// TIA Portal V19 export
FUNCTION_BLOCK "HOT_SKIDS"   // FB19, LAD
{ S7_Optimized_Access := 'TRUE' }
// stored: MemoryReserve 100, SetENOAutomatically false
   VAR_INPUT
      TEMP_SP : Real;
      AUTO : Bool;
      START : Bool;
      STOP : Bool;
      PUMP_SEL_1 : Bool;
      PUMP_SEL_2 : Bool;
      PUMP_SEL_3 : Bool;
      EMG : Bool;
      FS_HE_OUTLET : Bool;
      MGLT_LSP : Real;
      HOLD_RESUME : Bool;
      TT01_fault : Bool;
      TT02_fault : Bool;
      TT03_fault : Bool;
      TT04_fault : Bool;
      MGLT_FAULT : Bool;
      HEADER_PRESSURE_SP : Real;
      MGLT_PV : Real;
      TEMP_PV : Real;
      HEADER_PRESSURE_PV : Real;
      "PUMP 1RPM" : Real;
      "PUMP 1 RPM_SP" : Real;
      "PUMP 2 RPM" : Real;
      "PUMP 2 RPM_SP" : Real;
      "PUMP 3 RPM" : Real;
      "PUMP 3 RPM_SP" : Real;
   END_VAR
   VAR_OUTPUT
      PUMP_1_CMD : Bool;
      PUMP_2_CMD : Bool;
      PUMP_3_CMD : Bool;
      RUNNING : Bool;
      HS_CV_CMD : Bool;
      PUMP_SEL : Int;
      PUMP_1_FAULTY : Bool;
      PUMP_2_FAULTY : Bool;
      PUMP_3_FAULTY : Bool;
   END_VAR
   VAR
      "STEP" : Int;
      IEC_Timer_0_Instance { S7_SetPoint := 'True'} : TP_TIME;
      ALL_OK : Bool;
      TRIG_1 : Bool;
      TRIG_2 : Bool;
      TRIG_3 : Bool;
      TRIG_4 : Bool;
      TRIG_5 : Bool;
      TRIG_6 : Bool;
      TRIG_7 : Bool;
      IEC_Timer_0_Instance_1 { S7_SetPoint := 'True'} : TP_TIME;
      IEC_Timer_0_Instance_2 { S7_SetPoint := 'True'} : TP_TIME;
   END_VAR
   VAR_TEMP   // added for the SCL form of the ladder/FBD networks
      _w1 : Bool;
      _w2 : Bool;
      _w3 : Bool;
      _w4 : Bool;
   END_VAR
BEGIN

REGION Network 1: PRECHECK
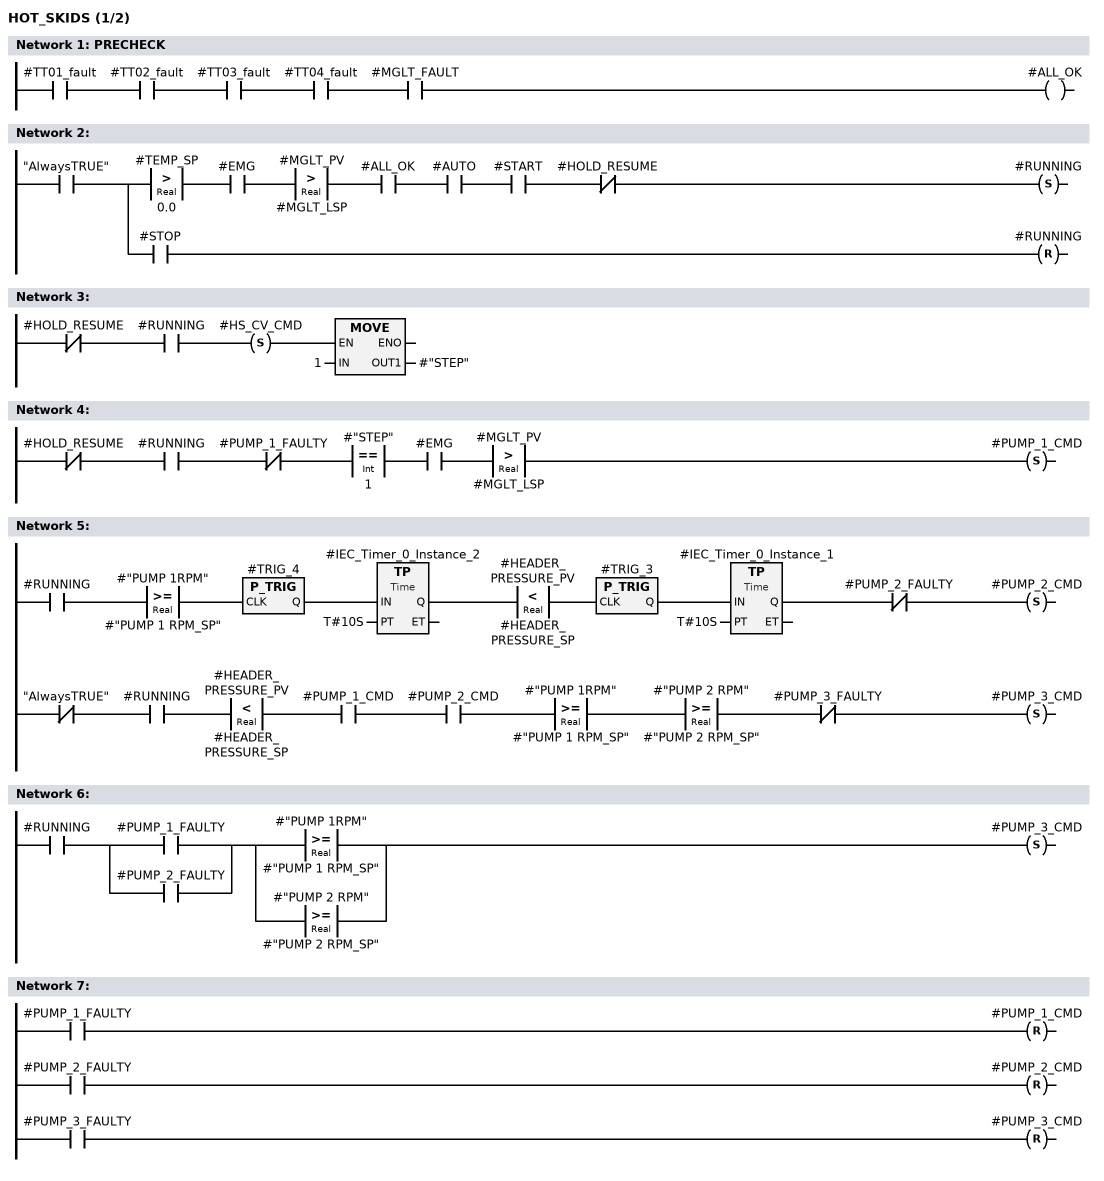
   RUNG wire#powerrail
      Contact( #TT01_fault )
      Contact( #TT02_fault )
      Contact( #TT03_fault )
      Contact( #TT04_fault )
      Contact( #MGLT_FAULT )
      Coil( #ALL_OK )
   END_RUNG
   // the same network as SCL:
   #ALL_OK := #TT01_fault AND #TT02_fault AND #TT03_fault AND #TT04_fault AND #MGLT_FAULT;
END_REGION

REGION Network 2
   RUNG wire#powerrail
      Contact( "AlwaysTRUE" )
      wire#w1
      { S7_Templates := "SrcType := Real" } GT_Contact(in1 := #TEMP_SP, in2 := 0.0)
      Contact( #EMG )
      { S7_Templates := "SrcType := Real" } GT_Contact(in1 := #MGLT_PV, in2 := #MGLT_LSP)
      Contact( #ALL_OK )
      Contact( #AUTO )
      Contact( #START )
      I_Contact( #HOLD_RESUME )
      S_Coil( #RUNNING )
   END_RUNG
   RUNG wire#w1
      Contact( #STOP )
      R_Coil( #RUNNING )
   END_RUNG
   // the same network as SCL:
   IF "AlwaysTRUE" AND (#TEMP_SP > 0.0) AND #EMG AND (#MGLT_PV > #MGLT_LSP) AND #ALL_OK AND #AUTO AND #START AND NOT #HOLD_RESUME THEN
       #RUNNING := TRUE;
   END_IF;
   IF "AlwaysTRUE" AND #STOP THEN #RUNNING := FALSE; END_IF;
END_REGION

REGION Network 3
   RUNG wire#powerrail
      I_Contact( #HOLD_RESUME )
      Contact( #RUNNING )
      S_Coil( #HS_CV_CMD )
      Move(in := 1, out1 => #"STEP")
   END_RUNG
   // the same network as SCL:
   IF NOT #HOLD_RESUME AND #RUNNING THEN
       #HS_CV_CMD := TRUE;
       #"STEP" := 1;
   END_IF;
END_REGION

REGION Network 4
   RUNG wire#powerrail
      I_Contact( #HOLD_RESUME )
      Contact( #RUNNING )
      I_Contact( #PUMP_1_FAULTY )
      { S7_Templates := "SrcType := Int" } EQ_Contact(in1 := #"STEP", in2 := 1)
      Contact( #EMG )
      { S7_Templates := "SrcType := Real" } GT_Contact(in1 := #MGLT_PV, in2 := #MGLT_LSP)
      S_Coil( #PUMP_1_CMD )
   END_RUNG
   // the same network as SCL:
   IF NOT #HOLD_RESUME AND #RUNNING AND NOT #PUMP_1_FAULTY AND (#"STEP" = 1) AND #EMG AND (#MGLT_PV > #MGLT_LSP) THEN
       #PUMP_1_CMD := TRUE;
   END_IF;
END_REGION

REGION Network 5
   RUNG wire#powerrail
      Contact( #RUNNING )
      { S7_Templates := "SrcType := Real" } GE_Contact(in1 := #"PUMP 1RPM", in2 := #"PUMP 1 RPM_SP")
      P_Trig( #TRIG_4 )
      { S7_Templates := "time_type := Time" } #IEC_Timer_0_Instance_2.TP(pt := T#10S, et =>)
      { S7_Templates := "SrcType := Real" } LT_Contact(in1 := #HEADER_PRESSURE_PV, in2 := #HEADER_PRESSURE_SP)
      P_Trig( #TRIG_3 )
      { S7_Templates := "time_type := Time" } #IEC_Timer_0_Instance_1.TP(pt := T#10S, et =>)
      I_Contact( #PUMP_2_FAULTY )
      S_Coil( #PUMP_2_CMD )
   END_RUNG
   RUNG wire#powerrail
      I_Contact( "AlwaysTRUE" )
      Contact( #RUNNING )
      { S7_Templates := "SrcType := Real" } LT_Contact(in1 := #HEADER_PRESSURE_PV, in2 := #HEADER_PRESSURE_SP)
      Contact( #PUMP_1_CMD )
      Contact( #PUMP_2_CMD )
      { S7_Templates := "SrcType := Real" } GE_Contact(in1 := #"PUMP 1RPM", in2 := #"PUMP 1 RPM_SP")
      { S7_Templates := "SrcType := Real" } GE_Contact(in1 := #"PUMP 2 RPM", in2 := #"PUMP 2 RPM_SP")
      I_Contact( #PUMP_3_FAULTY )
      S_Coil( #PUMP_3_CMD )
   END_RUNG
   // the same network as SCL:
   #_w1 := #RUNNING AND (#"PUMP 1RPM" >= #"PUMP 1 RPM_SP");
   #_w2 := #_w1 AND NOT #TRIG_4;   // rising edge
   #TRIG_4 := #_w1;
   #IEC_Timer_0_Instance_2(IN := #_w2, PT := T#10S);   // TP
   #_w3 := #IEC_Timer_0_Instance_2.Q AND (#HEADER_PRESSURE_PV < #HEADER_PRESSURE_SP);
   #_w4 := #_w3 AND NOT #TRIG_3;   // rising edge
   #TRIG_3 := #_w3;
   #IEC_Timer_0_Instance_1(IN := #_w4, PT := T#10S);   // TP
   IF #IEC_Timer_0_Instance_1.Q AND NOT #PUMP_2_FAULTY THEN #PUMP_2_CMD := TRUE; END_IF;
   IF NOT "AlwaysTRUE" AND #RUNNING AND (#HEADER_PRESSURE_PV < #HEADER_PRESSURE_SP) AND #PUMP_1_CMD AND #PUMP_2_CMD AND (#"PUMP 1RPM" >= #"PUMP 1 RPM_SP") AND (#"PUMP 2 RPM" >= #"PUMP 2 RPM_SP") AND NOT #PUMP_3_FAULTY THEN
       #PUMP_3_CMD := TRUE;
   END_IF;
END_REGION

REGION Network 6
   RUNG wire#powerrail
      Contact( #RUNNING )
      wire#w1
      Contact( #PUMP_1_FAULTY )
      wire#w2
      { S7_Templates := "SrcType := Real" } GE_Contact(in1 := #"PUMP 1RPM", in2 := #"PUMP 1 RPM_SP")
      wire#w3
      S_Coil( #PUMP_3_CMD )
   END_RUNG
   RUNG wire#w1
      Contact( #PUMP_2_FAULTY )
   END_RUNG wire#w2
   RUNG wire#w2
      { S7_Templates := "SrcType := Real" } GE_Contact(in1 := #"PUMP 2 RPM", in2 := #"PUMP 2 RPM_SP")
   END_RUNG wire#w3
   // the same network as SCL:
   IF #RUNNING AND (#PUMP_1_FAULTY OR #PUMP_2_FAULTY) AND ((#"PUMP 1RPM" >= #"PUMP 1 RPM_SP") OR (#"PUMP 2 RPM" >= #"PUMP 2 RPM_SP")) THEN
       #PUMP_3_CMD := TRUE;
   END_IF;
END_REGION

REGION Network 7
   RUNG wire#powerrail
      Contact( #PUMP_1_FAULTY )
      R_Coil( #PUMP_1_CMD )
   END_RUNG
   RUNG wire#powerrail
      Contact( #PUMP_2_FAULTY )
      R_Coil( #PUMP_2_CMD )
   END_RUNG
   RUNG wire#powerrail
      Contact( #PUMP_3_FAULTY )
      R_Coil( #PUMP_3_CMD )
   END_RUNG
   // the same network as SCL:
   IF #PUMP_1_FAULTY THEN #PUMP_1_CMD := FALSE; END_IF;
   IF #PUMP_2_FAULTY THEN #PUMP_2_CMD := FALSE; END_IF;
   IF #PUMP_3_FAULTY THEN #PUMP_3_CMD := FALSE; END_IF;
END_REGION

REGION Network 8
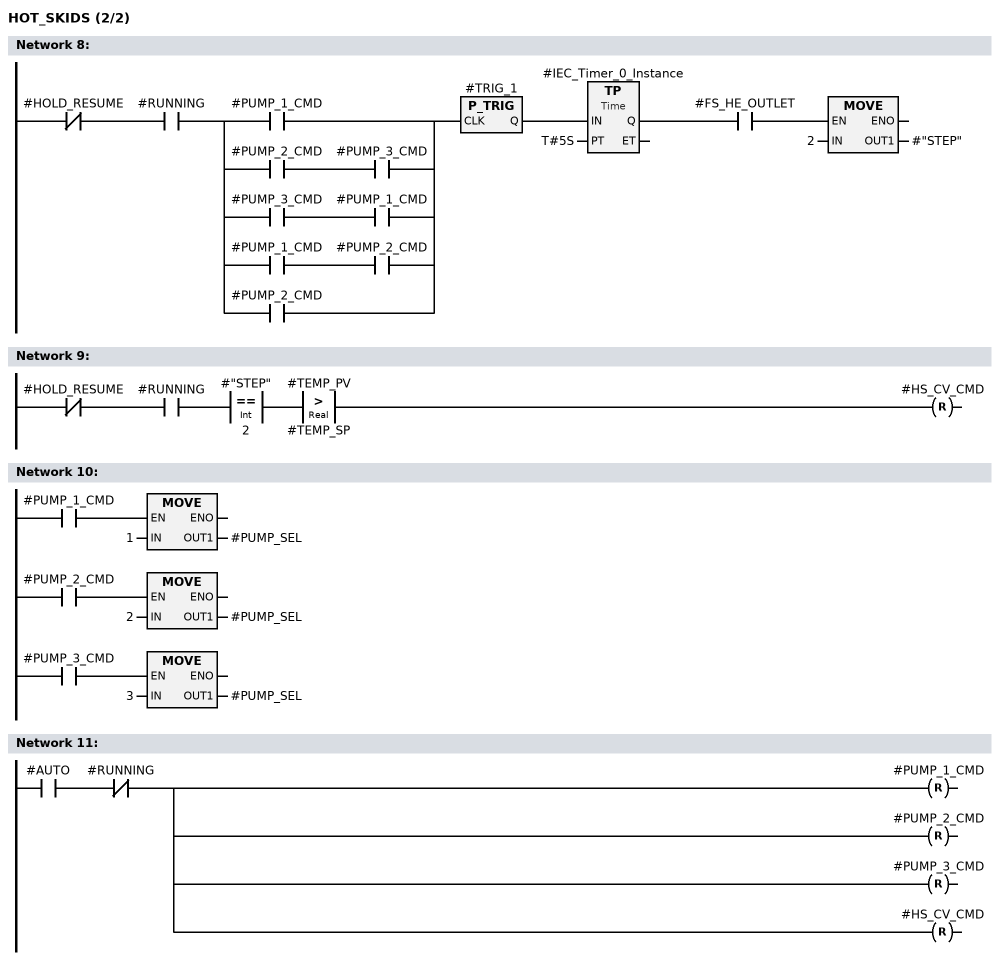
   RUNG wire#powerrail
      I_Contact( #HOLD_RESUME )
      Contact( #RUNNING )
      wire#w1
      Contact( #PUMP_1_CMD )
      wire#w2
      P_Trig( #TRIG_1 )
      { S7_Templates := "time_type := Time" } #IEC_Timer_0_Instance.TP(pt := T#5S, et =>)
      Contact( #FS_HE_OUTLET )
      Move(in := 2, out1 => #"STEP")
   END_RUNG
   RUNG wire#w1
      Contact( #PUMP_2_CMD )
      Contact( #PUMP_3_CMD )
   END_RUNG wire#w2
   RUNG wire#w1
      Contact( #PUMP_3_CMD )
      Contact( #PUMP_1_CMD )
   END_RUNG wire#w2
   RUNG wire#w1
      Contact( #PUMP_1_CMD )
      Contact( #PUMP_2_CMD )
   END_RUNG wire#w2
   RUNG wire#w1
      Contact( #PUMP_2_CMD )
   END_RUNG wire#w2
   // the same network as SCL:
   #_w1 := NOT #HOLD_RESUME AND #RUNNING AND (#PUMP_1_CMD OR (#PUMP_2_CMD AND #PUMP_3_CMD) OR (#PUMP_3_CMD AND #PUMP_1_CMD) OR (#PUMP_1_CMD AND #PUMP_2_CMD) OR #PUMP_2_CMD);
   #_w2 := #_w1 AND NOT #TRIG_1;   // rising edge
   #TRIG_1 := #_w1;
   #IEC_Timer_0_Instance(IN := #_w2, PT := T#5S);   // TP
   IF #IEC_Timer_0_Instance.Q AND #FS_HE_OUTLET THEN #"STEP" := 2; END_IF;
END_REGION

REGION Network 9
   RUNG wire#powerrail
      I_Contact( #HOLD_RESUME )
      Contact( #RUNNING )
      { S7_Templates := "SrcType := Int" } EQ_Contact(in1 := #"STEP", in2 := 2)
      { S7_Templates := "SrcType := Real" } GT_Contact(in1 := #TEMP_PV, in2 := #TEMP_SP)
      R_Coil( #HS_CV_CMD )
   END_RUNG
   // the same network as SCL:
   IF NOT #HOLD_RESUME AND #RUNNING AND (#"STEP" = 2) AND (#TEMP_PV > #TEMP_SP) THEN
       #HS_CV_CMD := FALSE;
   END_IF;
END_REGION

REGION Network 10
   RUNG wire#powerrail
      Contact( #PUMP_1_CMD )
      Move(in := 1, out1 => #PUMP_SEL)
   END_RUNG
   RUNG wire#powerrail
      Contact( #PUMP_2_CMD )
      Move(in := 2, out1 => #PUMP_SEL)
   END_RUNG
   RUNG wire#powerrail
      Contact( #PUMP_3_CMD )
      Move(in := 3, out1 => #PUMP_SEL)
   END_RUNG
   // the same network as SCL:
   IF #PUMP_1_CMD THEN #PUMP_SEL := 1; END_IF;
   IF #PUMP_2_CMD THEN #PUMP_SEL := 2; END_IF;
   IF #PUMP_3_CMD THEN #PUMP_SEL := 3; END_IF;
END_REGION

REGION Network 11
   RUNG wire#powerrail
      Contact( #AUTO )
      I_Contact( #RUNNING )
      wire#w1
      R_Coil( #PUMP_1_CMD )
   END_RUNG
   RUNG wire#w1
      R_Coil( #PUMP_2_CMD )
   END_RUNG
   RUNG wire#w1
      R_Coil( #PUMP_3_CMD )
   END_RUNG
   RUNG wire#w1
      R_Coil( #HS_CV_CMD )
   END_RUNG
   // the same network as SCL:
   IF #AUTO AND NOT #RUNNING THEN
       #PUMP_1_CMD := FALSE;
       #PUMP_2_CMD := FALSE;
       #PUMP_3_CMD := FALSE;
       #HS_CV_CMD := FALSE;
   END_IF;
END_REGION
END_FUNCTION_BLOCK
